DATA_BLOCK "CallerData"
{ S7_Optimized_Access := 'TRUE' }
VERSION : 0.1
NON_RETAIN
"Caller"

BEGIN

END_DATA_BLOCK

